SYSTEM FU_Demo
  (* Version 1.0, 2026-11-02, Franz Höpfinger *)
  IMPORT FBs::FU_Demo::FU_Demo_Konstanten::APIXON;
  APPLICATION FU_DemoApp
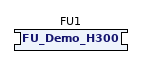
    SUBAPPS
      FU1 : FBs::FU_Demo::FU_Demo_H300;
    END_SUBAPPS
  END_APPLICATION
  DEVICE APIXON : iec61499::system::FORTE_PC(MGR_ID := APIXON (* Device manager socket ID *))
    {SET_ATTRIBUTE(Profile, HOLOBLOC)}
    RESOURCE EMB_RES : iec61499::system::EMB_RES
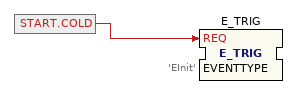
      FBS
        E_TRIG : iec61499::events::E_TRIG(EVENTTYPE := 'EInit');
      END_FBS
      EVENT_CONNECTIONS
        START.COLD TO E_TRIG.REQ;
      END_CONNECTIONS
    END_RESOURCE
  END_DEVICE
  MAPPINGS
    FU_DemoApp.FU1 ON APIXON.EMB_RES;
  END_MAPPINGS
  SEGMENTS
    Ethernet : iec61499::system::Ethernet;
  END_SEGMENTS
  LINKS
    APIXON => Ethernet;
  END_LINKS
END_SYSTEM
